Fanuc KAREL source: kd00037.KL

-- PROVISIONAL review KL for V1013-1; original PC SHA256 340f200e0b70047e08b8e89d0cf1a292fd413fd2284839e5aa22f7e74d58e6ac
-- Incomplete behavior may be omitted. Consult companion uncertainty JSON. Do not deploy.
PROGRAM KD00037
%NOLOCKGROUP
VAR
  I : INTEGER
  J : INTEGER
  B : BOOLEAN
  R : REAL
  S : STRING[80]
BEGIN
  -- UNRESOLVED_PC offsets 5-18; opcodes 9D,81,18,9D,1B,9D,12,9C,13,04
  -- UNRESOLVED_PC offsets 23-27; opcodes 7F
END KD00037
